(* IEC 61131-3 sources: STAR-PLC-Agent/results/raw/pilot_pair_2026-11-10T143217961073+0000/PUB001_star/sim_00, 1 file *)

(* ---- test_program.st ---- *)
PROGRAM PLC_PRG
VAR
 BenchStep : UDINT := 0;
 BenchCalls : UDINT := 0;
 BenchDone : BOOL := FALSE;
 BenchUut0 : FB_Task;
 BenchUut1 : FB_Task;
 TraceIn_bottleSensor : ARRAY[0..12] OF BOOL;
 TraceIn_cleaningConfirmButton : ARRAY[0..12] OF BOOL;
 TraceIn_fillingConfirmButton : ARRAY[0..12] OF BOOL;
 TraceIn_cappingConfirmButton : ARRAY[0..12] OF BOOL;
 TraceIn_packingConfirmButton : ARRAY[0..12] OF BOOL;
 TraceIn_finishedButton : ARRAY[0..12] OF BOOL;
 TraceOut_Pump_Motor : ARRAY[0..12] OF BOOL;
 TraceOut_Filling_Valve : ARRAY[0..12] OF BOOL;
 TraceOut_Capping_Machine : ARRAY[0..12] OF BOOL;
 TraceOut_Packing_Machine : ARRAY[0..12] OF BOOL;
 TraceOut_Completion_Light : ARRAY[0..12] OF BOOL;
END_VAR

IF NOT BenchDone THEN
 CASE BenchStep OF
 0:
   BenchUut0.bottleSensor := TRUE;
   BenchUut0.cleaningConfirmButton := FALSE;
   BenchUut0.fillingConfirmButton := FALSE;
   BenchUut0.cappingConfirmButton := FALSE;
   BenchUut0.packingConfirmButton := FALSE;
   BenchUut0.finishedButton := FALSE;
   TraceIn_bottleSensor[0] := BenchUut0.bottleSensor;
   TraceIn_cleaningConfirmButton[0] := BenchUut0.cleaningConfirmButton;
   TraceIn_fillingConfirmButton[0] := BenchUut0.fillingConfirmButton;
   TraceIn_cappingConfirmButton[0] := BenchUut0.cappingConfirmButton;
   TraceIn_packingConfirmButton[0] := BenchUut0.packingConfirmButton;
   TraceIn_finishedButton[0] := BenchUut0.finishedButton;
   BenchUut0();
   TraceOut_Pump_Motor[0] := BenchUut0.Pump_Motor;
   TraceOut_Filling_Valve[0] := BenchUut0.Filling_Valve;
   TraceOut_Capping_Machine[0] := BenchUut0.Capping_Machine;
   TraceOut_Packing_Machine[0] := BenchUut0.Packing_Machine;
   TraceOut_Completion_Light[0] := BenchUut0.Completion_Light;
   BenchCalls := BenchCalls + 1;
 1:
   BenchUut0.bottleSensor := FALSE;
   BenchUut0.cleaningConfirmButton := TRUE;
   BenchUut0.fillingConfirmButton := FALSE;
   BenchUut0.cappingConfirmButton := FALSE;
   BenchUut0.packingConfirmButton := FALSE;
   BenchUut0.finishedButton := FALSE;
   TraceIn_bottleSensor[1] := BenchUut0.bottleSensor;
   TraceIn_cleaningConfirmButton[1] := BenchUut0.cleaningConfirmButton;
   TraceIn_fillingConfirmButton[1] := BenchUut0.fillingConfirmButton;
   TraceIn_cappingConfirmButton[1] := BenchUut0.cappingConfirmButton;
   TraceIn_packingConfirmButton[1] := BenchUut0.packingConfirmButton;
   TraceIn_finishedButton[1] := BenchUut0.finishedButton;
   BenchUut0();
   TraceOut_Pump_Motor[1] := BenchUut0.Pump_Motor;
   TraceOut_Filling_Valve[1] := BenchUut0.Filling_Valve;
   TraceOut_Capping_Machine[1] := BenchUut0.Capping_Machine;
   TraceOut_Packing_Machine[1] := BenchUut0.Packing_Machine;
   TraceOut_Completion_Light[1] := BenchUut0.Completion_Light;
   BenchCalls := BenchCalls + 1;
 2:
   BenchUut0.bottleSensor := FALSE;
   BenchUut0.cleaningConfirmButton := FALSE;
   BenchUut0.fillingConfirmButton := TRUE;
   BenchUut0.cappingConfirmButton := FALSE;
   BenchUut0.packingConfirmButton := FALSE;
   BenchUut0.finishedButton := FALSE;
   TraceIn_bottleSensor[2] := BenchUut0.bottleSensor;
   TraceIn_cleaningConfirmButton[2] := BenchUut0.cleaningConfirmButton;
   TraceIn_fillingConfirmButton[2] := BenchUut0.fillingConfirmButton;
   TraceIn_cappingConfirmButton[2] := BenchUut0.cappingConfirmButton;
   TraceIn_packingConfirmButton[2] := BenchUut0.packingConfirmButton;
   TraceIn_finishedButton[2] := BenchUut0.finishedButton;
   BenchUut0();
   TraceOut_Pump_Motor[2] := BenchUut0.Pump_Motor;
   TraceOut_Filling_Valve[2] := BenchUut0.Filling_Valve;
   TraceOut_Capping_Machine[2] := BenchUut0.Capping_Machine;
   TraceOut_Packing_Machine[2] := BenchUut0.Packing_Machine;
   TraceOut_Completion_Light[2] := BenchUut0.Completion_Light;
   BenchCalls := BenchCalls + 1;
 3:
   BenchUut0.bottleSensor := FALSE;
   BenchUut0.cleaningConfirmButton := FALSE;
   BenchUut0.fillingConfirmButton := FALSE;
   BenchUut0.cappingConfirmButton := TRUE;
   BenchUut0.packingConfirmButton := FALSE;
   BenchUut0.finishedButton := FALSE;
   TraceIn_bottleSensor[3] := BenchUut0.bottleSensor;
   TraceIn_cleaningConfirmButton[3] := BenchUut0.cleaningConfirmButton;
   TraceIn_fillingConfirmButton[3] := BenchUut0.fillingConfirmButton;
   TraceIn_cappingConfirmButton[3] := BenchUut0.cappingConfirmButton;
   TraceIn_packingConfirmButton[3] := BenchUut0.packingConfirmButton;
   TraceIn_finishedButton[3] := BenchUut0.finishedButton;
   BenchUut0();
   TraceOut_Pump_Motor[3] := BenchUut0.Pump_Motor;
   TraceOut_Filling_Valve[3] := BenchUut0.Filling_Valve;
   TraceOut_Capping_Machine[3] := BenchUut0.Capping_Machine;
   TraceOut_Packing_Machine[3] := BenchUut0.Packing_Machine;
   TraceOut_Completion_Light[3] := BenchUut0.Completion_Light;
   BenchCalls := BenchCalls + 1;
 4:
   BenchUut0.bottleSensor := FALSE;
   BenchUut0.cleaningConfirmButton := FALSE;
   BenchUut0.fillingConfirmButton := FALSE;
   BenchUut0.cappingConfirmButton := FALSE;
   BenchUut0.packingConfirmButton := TRUE;
   BenchUut0.finishedButton := FALSE;
   TraceIn_bottleSensor[4] := BenchUut0.bottleSensor;
   TraceIn_cleaningConfirmButton[4] := BenchUut0.cleaningConfirmButton;
   TraceIn_fillingConfirmButton[4] := BenchUut0.fillingConfirmButton;
   TraceIn_cappingConfirmButton[4] := BenchUut0.cappingConfirmButton;
   TraceIn_packingConfirmButton[4] := BenchUut0.packingConfirmButton;
   TraceIn_finishedButton[4] := BenchUut0.finishedButton;
   BenchUut0();
   TraceOut_Pump_Motor[4] := BenchUut0.Pump_Motor;
   TraceOut_Filling_Valve[4] := BenchUut0.Filling_Valve;
   TraceOut_Capping_Machine[4] := BenchUut0.Capping_Machine;
   TraceOut_Packing_Machine[4] := BenchUut0.Packing_Machine;
   TraceOut_Completion_Light[4] := BenchUut0.Completion_Light;
   BenchCalls := BenchCalls + 1;
 5:
   BenchUut0.bottleSensor := FALSE;
   BenchUut0.cleaningConfirmButton := FALSE;
   BenchUut0.fillingConfirmButton := FALSE;
   BenchUut0.cappingConfirmButton := FALSE;
   BenchUut0.packingConfirmButton := FALSE;
   BenchUut0.finishedButton := TRUE;
   TraceIn_bottleSensor[5] := BenchUut0.bottleSensor;
   TraceIn_cleaningConfirmButton[5] := BenchUut0.cleaningConfirmButton;
   TraceIn_fillingConfirmButton[5] := BenchUut0.fillingConfirmButton;
   TraceIn_cappingConfirmButton[5] := BenchUut0.cappingConfirmButton;
   TraceIn_packingConfirmButton[5] := BenchUut0.packingConfirmButton;
   TraceIn_finishedButton[5] := BenchUut0.finishedButton;
   BenchUut0();
   TraceOut_Pump_Motor[5] := BenchUut0.Pump_Motor;
   TraceOut_Filling_Valve[5] := BenchUut0.Filling_Valve;
   TraceOut_Capping_Machine[5] := BenchUut0.Capping_Machine;
   TraceOut_Packing_Machine[5] := BenchUut0.Packing_Machine;
   TraceOut_Completion_Light[5] := BenchUut0.Completion_Light;
   BenchCalls := BenchCalls + 1;
 6:
   BenchUut1.bottleSensor := TRUE;
   BenchUut1.cleaningConfirmButton := FALSE;
   BenchUut1.fillingConfirmButton := TRUE;
   BenchUut1.cappingConfirmButton := FALSE;
   BenchUut1.packingConfirmButton := FALSE;
   BenchUut1.finishedButton := FALSE;
   TraceIn_bottleSensor[6] := BenchUut1.bottleSensor;
   TraceIn_cleaningConfirmButton[6] := BenchUut1.cleaningConfirmButton;
   TraceIn_fillingConfirmButton[6] := BenchUut1.fillingConfirmButton;
   TraceIn_cappingConfirmButton[6] := BenchUut1.cappingConfirmButton;
   TraceIn_packingConfirmButton[6] := BenchUut1.packingConfirmButton;
   TraceIn_finishedButton[6] := BenchUut1.finishedButton;
   BenchUut1();
   TraceOut_Pump_Motor[6] := BenchUut1.Pump_Motor;
   TraceOut_Filling_Valve[6] := BenchUut1.Filling_Valve;
   TraceOut_Capping_Machine[6] := BenchUut1.Capping_Machine;
   TraceOut_Packing_Machine[6] := BenchUut1.Packing_Machine;
   TraceOut_Completion_Light[6] := BenchUut1.Completion_Light;
   BenchCalls := BenchCalls + 1;
 7:
   BenchUut1.bottleSensor := FALSE;
   BenchUut1.cleaningConfirmButton := TRUE;
   BenchUut1.fillingConfirmButton := FALSE;
   BenchUut1.cappingConfirmButton := TRUE;
   BenchUut1.packingConfirmButton := FALSE;
   BenchUut1.finishedButton := FALSE;
   TraceIn_bottleSensor[7] := BenchUut1.bottleSensor;
   TraceIn_cleaningConfirmButton[7] := BenchUut1.cleaningConfirmButton;
   TraceIn_fillingConfirmButton[7] := BenchUut1.fillingConfirmButton;
   TraceIn_cappingConfirmButton[7] := BenchUut1.cappingConfirmButton;
   TraceIn_packingConfirmButton[7] := BenchUut1.packingConfirmButton;
   TraceIn_finishedButton[7] := BenchUut1.finishedButton;
   BenchUut1();
   TraceOut_Pump_Motor[7] := BenchUut1.Pump_Motor;
   TraceOut_Filling_Valve[7] := BenchUut1.Filling_Valve;
   TraceOut_Capping_Machine[7] := BenchUut1.Capping_Machine;
   TraceOut_Packing_Machine[7] := BenchUut1.Packing_Machine;
   TraceOut_Completion_Light[7] := BenchUut1.Completion_Light;
   BenchCalls := BenchCalls + 1;
 8:
   BenchUut1.bottleSensor := FALSE;
   BenchUut1.cleaningConfirmButton := FALSE;
   BenchUut1.fillingConfirmButton := TRUE;
   BenchUut1.cappingConfirmButton := FALSE;
   BenchUut1.packingConfirmButton := TRUE;
   BenchUut1.finishedButton := FALSE;
   TraceIn_bottleSensor[8] := BenchUut1.bottleSensor;
   TraceIn_cleaningConfirmButton[8] := BenchUut1.cleaningConfirmButton;
   TraceIn_fillingConfirmButton[8] := BenchUut1.fillingConfirmButton;
   TraceIn_cappingConfirmButton[8] := BenchUut1.cappingConfirmButton;
   TraceIn_packingConfirmButton[8] := BenchUut1.packingConfirmButton;
   TraceIn_finishedButton[8] := BenchUut1.finishedButton;
   BenchUut1();
   TraceOut_Pump_Motor[8] := BenchUut1.Pump_Motor;
   TraceOut_Filling_Valve[8] := BenchUut1.Filling_Valve;
   TraceOut_Capping_Machine[8] := BenchUut1.Capping_Machine;
   TraceOut_Packing_Machine[8] := BenchUut1.Packing_Machine;
   TraceOut_Completion_Light[8] := BenchUut1.Completion_Light;
   BenchCalls := BenchCalls + 1;
 9:
   BenchUut1.bottleSensor := FALSE;
   BenchUut1.cleaningConfirmButton := FALSE;
   BenchUut1.fillingConfirmButton := FALSE;
   BenchUut1.cappingConfirmButton := TRUE;
   BenchUut1.packingConfirmButton := FALSE;
   BenchUut1.finishedButton := TRUE;
   TraceIn_bottleSensor[9] := BenchUut1.bottleSensor;
   TraceIn_cleaningConfirmButton[9] := BenchUut1.cleaningConfirmButton;
   TraceIn_fillingConfirmButton[9] := BenchUut1.fillingConfirmButton;
   TraceIn_cappingConfirmButton[9] := BenchUut1.cappingConfirmButton;
   TraceIn_packingConfirmButton[9] := BenchUut1.packingConfirmButton;
   TraceIn_finishedButton[9] := BenchUut1.finishedButton;
   BenchUut1();
   TraceOut_Pump_Motor[9] := BenchUut1.Pump_Motor;
   TraceOut_Filling_Valve[9] := BenchUut1.Filling_Valve;
   TraceOut_Capping_Machine[9] := BenchUut1.Capping_Machine;
   TraceOut_Packing_Machine[9] := BenchUut1.Packing_Machine;
   TraceOut_Completion_Light[9] := BenchUut1.Completion_Light;
   BenchCalls := BenchCalls + 1;
 10:
   BenchUut1.bottleSensor := FALSE;
   BenchUut1.cleaningConfirmButton := FALSE;
   BenchUut1.fillingConfirmButton := FALSE;
   BenchUut1.cappingConfirmButton := FALSE;
   BenchUut1.packingConfirmButton := TRUE;
   BenchUut1.finishedButton := TRUE;
   TraceIn_bottleSensor[10] := BenchUut1.bottleSensor;
   TraceIn_cleaningConfirmButton[10] := BenchUut1.cleaningConfirmButton;
   TraceIn_fillingConfirmButton[10] := BenchUut1.fillingConfirmButton;
   TraceIn_cappingConfirmButton[10] := BenchUut1.cappingConfirmButton;
   TraceIn_packingConfirmButton[10] := BenchUut1.packingConfirmButton;
   TraceIn_finishedButton[10] := BenchUut1.finishedButton;
   BenchUut1();
   TraceOut_Pump_Motor[10] := BenchUut1.Pump_Motor;
   TraceOut_Filling_Valve[10] := BenchUut1.Filling_Valve;
   TraceOut_Capping_Machine[10] := BenchUut1.Capping_Machine;
   TraceOut_Packing_Machine[10] := BenchUut1.Packing_Machine;
   TraceOut_Completion_Light[10] := BenchUut1.Completion_Light;
   BenchCalls := BenchCalls + 1;
 11:
   BenchUut1.bottleSensor := TRUE;
   BenchUut1.cleaningConfirmButton := FALSE;
   BenchUut1.fillingConfirmButton := FALSE;
   BenchUut1.cappingConfirmButton := FALSE;
   BenchUut1.packingConfirmButton := FALSE;
   BenchUut1.finishedButton := TRUE;
   TraceIn_bottleSensor[11] := BenchUut1.bottleSensor;
   TraceIn_cleaningConfirmButton[11] := BenchUut1.cleaningConfirmButton;
   TraceIn_fillingConfirmButton[11] := BenchUut1.fillingConfirmButton;
   TraceIn_cappingConfirmButton[11] := BenchUut1.cappingConfirmButton;
   TraceIn_packingConfirmButton[11] := BenchUut1.packingConfirmButton;
   TraceIn_finishedButton[11] := BenchUut1.finishedButton;
   BenchUut1();
   TraceOut_Pump_Motor[11] := BenchUut1.Pump_Motor;
   TraceOut_Filling_Valve[11] := BenchUut1.Filling_Valve;
   TraceOut_Capping_Machine[11] := BenchUut1.Capping_Machine;
   TraceOut_Packing_Machine[11] := BenchUut1.Packing_Machine;
   TraceOut_Completion_Light[11] := BenchUut1.Completion_Light;
   BenchCalls := BenchCalls + 1;
 12:
   BenchUut1.bottleSensor := TRUE;
   BenchUut1.cleaningConfirmButton := FALSE;
   BenchUut1.fillingConfirmButton := FALSE;
   BenchUut1.cappingConfirmButton := FALSE;
   BenchUut1.packingConfirmButton := FALSE;
   BenchUut1.finishedButton := FALSE;
   TraceIn_bottleSensor[12] := BenchUut1.bottleSensor;
   TraceIn_cleaningConfirmButton[12] := BenchUut1.cleaningConfirmButton;
   TraceIn_fillingConfirmButton[12] := BenchUut1.fillingConfirmButton;
   TraceIn_cappingConfirmButton[12] := BenchUut1.cappingConfirmButton;
   TraceIn_packingConfirmButton[12] := BenchUut1.packingConfirmButton;
   TraceIn_finishedButton[12] := BenchUut1.finishedButton;
   BenchUut1();
   TraceOut_Pump_Motor[12] := BenchUut1.Pump_Motor;
   TraceOut_Filling_Valve[12] := BenchUut1.Filling_Valve;
   TraceOut_Capping_Machine[12] := BenchUut1.Capping_Machine;
   TraceOut_Packing_Machine[12] := BenchUut1.Packing_Machine;
   TraceOut_Completion_Light[12] := BenchUut1.Completion_Light;
   BenchCalls := BenchCalls + 1;
 END_CASE;
 BenchStep := BenchStep + 1;
 IF BenchStep >= 13 THEN BenchDone := TRUE; END_IF;
END_IF;
END_PROGRAM
